Fanuc KAREL source: kb00158.KL

PROGRAM KB00158
%STACKSIZE=65535
%PRIORITY=65535
%NOLOCKGROUP
VAR
P1 : INTEGER
P2 : INTEGER
BEGIN
P1=1
P2=1
SEND_EVENTPC(P1,P2)
END KB00158
